TYPE ST_AlarmHistoryEntry :
STRUCT
    sMessageText : STRING(255);
    nTimestamp   : ULINT;
    eSeverity    : TcEventSeverity;
END_STRUCT
END_TYPE

(* stored: Version 1.1.0.1, ProductVersion 3.1.4024.15
   DUT ST_AlarmHistoryEntry: Id {6f97cb22-27a0-494c-bce9-8dc9e0a0ec6a} *)
